# EPICS substitutions: db/Beckhoff_7XXX/ecmcEX72XX_OPT_encoder.substitutions
file "ecmcEL72XX_ENC.template"
{
  pattern {CH_ID}
          {"$(OPT_CH_ID=01)"}
}
